// Generated by voz_llm_plc_agent
// Target: Siemens TIA Portal V18 - SCL external source
// Review and compile before any download to physical hardware.

FUNCTION_BLOCK "PLC_PRG"
{ S7_Optimized_Access := 'TRUE' }
VERSION : 0.1
VAR_INPUT
   I_Start : Bool := FALSE;
   I_Emergency : Bool := FALSE;
END_VAR
VAR_OUTPUT
   Q_Lamp : Bool := FALSE;
END_VAR
BEGIN
(* Salida directa habilitada por entrada *)
#Q_Lamp := #I_Start AND NOT #I_Emergency;
(* Bloqueo: #I_Emergency fuerza a FALSE #Q_Lamp de inmediato *)
IF #I_Emergency THEN
    #Q_Lamp := FALSE;
END_IF;
END_FUNCTION_BLOCK

DATA_BLOCK "DB_PLC_PRG"
{ S7_Optimized_Access := 'TRUE' }
VERSION : 0.1
NON_RETAIN
"PLC_PRG"
BEGIN
END_DATA_BLOCK

ORGANIZATION_BLOCK "Main"
{ S7_Optimized_Access := 'TRUE' }
VERSION : 0.1
BEGIN
   "DB_PLC_PRG"(
      I_Start := "I_Start",
      I_Emergency := "I_Emergency",
      Q_Lamp => "Q_Lamp"
   );
END_ORGANIZATION_BLOCK
